(* IEC 61131-3 sources: plc-vscode/tests/st/test-ready/trust-platform/examples/OSCAT/solar_lighting_clock/non-oop/src, 3 files *)

(* ---- Configuration.st ---- *)
CONFIGURATION SolarLightingClockClassicConfiguration
RESOURCE Cpu0 ON PLC
    TASK MainTask (INTERVAL := T#1s, PRIORITY := 1);
    PROGRAM Main WITH MainTask : Main;
END_RESOURCE
END_CONFIGURATION

(* ---- Main.st ---- *)
PROGRAM Main
VAR
    ConstantsReady : BOOL;
    CalendarData : CALENDAR;
    Holidays : ARRAY[0..29] OF HOLIDAY_DATA;
    CalendarCalculator : CALENDAR_CALC;
    ExteriorLightingRequest : BOOL;
    LocalYear : INT;
END_VAR

ConstantsReady := OSCAT_BASIC_Constants();
CalendarData.UTC := DT#2026-04-26-10:00:00;
CalendarData.DST_EN := TRUE;
CalendarData.OFFSET := INT#60;
CalendarData.LANGUAGE := INT#1;
CalendarData.LATITUDE := REAL#59.3293;
CalendarData.LONGITUDE := REAL#18.0686;
CalendarCalculator(SPE := TRUE, H := REAL#-0.8333333, XCAL := CalendarData, HOLIDAYS := Holidays);
ExteriorLightingRequest := CalendarData.NIGHT;
LocalYear := CalendarData.YEAR;
END_PROGRAM

(* ---- Tests.st ---- *)
TEST_PROGRAM SolarLightingClockClassicCalculatesLocalCalendar
VAR
    ConstantsReady : BOOL;
    CalendarData : CALENDAR;
    Holidays : ARRAY[0..29] OF HOLIDAY_DATA;
    CalendarCalculator : CALENDAR_CALC;
END_VAR

ConstantsReady := OSCAT_BASIC_Constants();
CalendarData.UTC := DT#2026-04-26-10:00:00;
CalendarData.DST_EN := TRUE;
CalendarData.OFFSET := INT#60;
CalendarData.LANGUAGE := INT#1;
CalendarData.LATITUDE := REAL#59.3293;
CalendarData.LONGITUDE := REAL#18.0686;
CalendarCalculator(SPE := TRUE, H := REAL#-0.8333333, XCAL := CalendarData, HOLIDAYS := Holidays);

ASSERT_TRUE(IN := ConstantsReady);
ASSERT_EQUAL(EXPECTED := INT#2026, ACTUAL := CalendarData.YEAR);
ASSERT_EQUAL(EXPECTED := INT#4, ACTUAL := CalendarData.MONTH);
ASSERT_EQUAL(EXPECTED := INT#26, ACTUAL := CalendarData.DAY);
END_TEST_PROGRAM
